Staubli VAL3: Action.pjx

--- Action.pjx ---
Parameters version=s8.10.3Cs9_BS2093 stackSize=5000 millimeterUnit=true
Program file=_tActCtrl.pgx
Program file=action.pgx
Program file=action_do.pgx
Program file=addActCmd.pgx
Program file=checkMoveId.pgx
Program file=clearActStack.pgx
Program file=create.pgx
Program file=init.pgx
Program file=kill.pgx
Program file=moveJToJoint.pgx
Program file=moveLJToPoint.pgx
Program file=pushActCmd.pgx
Program file=removeActCmd.pgx
Program file=resetMoveId.pgx
Program file=start.pgx
Program file=stop.pgx
Data file=Action.dtx
Library alias=io path=Disk://source/projectSource/io/io.pjx
Library alias=rs path=Disk://source/projectSource/robotStatus/robotStatus.pjx
Library alias=actionData path=Disk://data/actionData/actionData.pjx
Type name=actionIO path=Disk://source/template/action/action.pjx
Type name=actCmdType path=Disk://source/template/actCmd/actCmd.pjx

--- Action.dtx ---
actCmdType actCmd[40]
  [0]
    bool bActFinish
    num nActionID
    num nMoveID
    string sActName
  [1]
    bool bActFinish
    num nActionID
    num nMoveID
    string sActName
  [2]
    bool bActFinish
    num nActionID
    num nMoveID
    string sActName
  [3]
    bool bActFinish
    num nActionID
    num nMoveID
    string sActName
  [4]
    bool bActFinish
    num nActionID
    num nMoveID
    string sActName
  [5]
    bool bActFinish
    num nActionID
    num nMoveID
    string sActName
  [6]
    bool bActFinish
    num nActionID
    num nMoveID
    string sActName
  [7]
    bool bActFinish
    num nActionID
    num nMoveID
    string sActName
  [8]
    bool bActFinish
    num nActionID
    num nMoveID
    string sActName
  [9]
    bool bActFinish
    num nActionID
    num nMoveID
    string sActName
  [10]
    bool bActFinish
    num nActionID
    num nMoveID
    string sActName
  [11]
    bool bActFinish
    num nActionID
    num nMoveID
    string sActName
  [12]
    bool bActFinish
    num nActionID
    num nMoveID
    string sActName
  [13]
    bool bActFinish
    num nActionID
    num nMoveID
    string sActName
  [14]
    bool bActFinish
    num nActionID
    num nMoveID
    string sActName
  [15]
    bool bActFinish
    num nActionID
    num nMoveID
    string sActName
  [16]
    bool bActFinish
    num nActionID
    num nMoveID
    string sActName
  [17]
    bool bActFinish
    num nActionID
    num nMoveID
    string sActName
  [18]
    bool bActFinish
    num nActionID
    num nMoveID
    string sActName
  [19]
    bool bActFinish
    num nActionID
    num nMoveID
    string sActName
  [20]
    bool bActFinish
    num nActionID
    num nMoveID
    string sActName
  [21]
    bool bActFinish
    num nActionID
    num nMoveID
    string sActName
  [22]
    bool bActFinish
    num nActionID
    num nMoveID
    string sActName
  [23]
    bool bActFinish
    num nActionID
    num nMoveID
    string sActName
  [24]
    bool bActFinish
    num nActionID
    num nMoveID
    string sActName
  [25]
    bool bActFinish
    num nActionID
    num nMoveID
    string sActName
  [26]
    bool bActFinish
    num nActionID
    num nMoveID
    string sActName
  [27]
    bool bActFinish
    num nActionID
    num nMoveID
    string sActName
  [28]
    bool bActFinish
    num nActionID
    num nMoveID
    string sActName
  [29]
    bool bActFinish
    num nActionID
    num nMoveID
    string sActName
  [30]
    bool bActFinish
    num nActionID
    num nMoveID
    string sActName
  [31]
    bool bActFinish
    num nActionID
    num nMoveID
    string sActName
  [32]
    bool bActFinish
    num nActionID
    num nMoveID
    string sActName
  [33]
    bool bActFinish
    num nActionID
    num nMoveID
    string sActName
  [34]
    bool bActFinish
    num nActionID
    num nMoveID
    string sActName
  [35]
    bool bActFinish
    num nActionID
    num nMoveID
    string sActName
  [36]
    bool bActFinish
    num nActionID
    num nMoveID
    string sActName
  [37]
    bool bActFinish
    num nActionID
    num nMoveID
    string sActName
  [38]
    bool bActFinish
    num nActionID
    num nMoveID
    string sActName
  [39]
    bool bActFinish
    num nActionID
    num nMoveID
    string sActName
actionIO aActionUsing
  [0]
    num nActIO
    num nActResult
    num nActType
actionIO actPrt[40]
  [0]
    num nActIO
    num nActResult
    num nActType
  [1]
    num nActIO
    num nActResult
    num nActType
  [2]
    num nActIO
    num nActResult
    num nActType
  [3]
    num nActIO
    num nActResult
    num nActType
  [4]
    num nActIO
    num nActResult
    num nActType
  [5]
    num nActIO
    num nActResult
    num nActType
  [6]
    num nActIO
    num nActResult
    num nActType
  [7]
    num nActIO
    num nActResult
    num nActType
  [8]
    num nActIO
    num nActResult
    num nActType
  [9]
    num nActIO
    num nActResult
    num nActType
  [10]
    num nActIO
    num nActResult
    num nActType
  [11]
    num nActIO
    num nActResult
    num nActType
  [12]
    num nActIO
    num nActResult
    num nActType
  [13]
    num nActIO
    num nActResult
    num nActType
  [14]
    num nActIO
    num nActResult
    num nActType
  [15]
    num nActIO
    num nActResult
    num nActType
  [16]
    num nActIO
    num nActResult
    num nActType
  [17]
    num nActIO
    num nActResult
    num nActType
  [18]
    num nActIO
    num nActResult
    num nActType
  [19]
    num nActIO
    num nActResult
    num nActType
  [20]
    num nActIO
    num nActResult
    num nActType
  [21]
    num nActIO
    num nActResult
    num nActType
  [22]
    num nActIO
    num nActResult
    num nActType
  [23]
    num nActIO
    num nActResult
    num nActType
  [24]
    num nActIO
    num nActResult
    num nActType
  [25]
    num nActIO
    num nActResult
    num nActType
  [26]
    num nActIO
    num nActResult
    num nActType
  [27]
    num nActIO
    num nActResult
    num nActType
  [28]
    num nActIO
    num nActResult
    num nActType
  [29]
    num nActIO
    num nActResult
    num nActType
  [30]
    num nActIO
    num nActResult
    num nActType
  [31]
    num nActIO
    num nActResult
    num nActType
  [32]
    num nActIO
    num nActResult
    num nActType
  [33]
    num nActIO
    num nActResult
    num nActType
  [34]
    num nActIO
    num nActResult
    num nActType
  [35]
    num nActIO
    num nActResult
    num nActType
  [36]
    num nActIO
    num nActResult
    num nActType
  [37]
    num nActIO
    num nActResult
    num nActType
  [38]
    num nActIO
    num nActResult
    num nActType
  [39]
    num nActIO
    num nActResult
    num nActType
bool bPushToStack
public num _nActStackIndex
num _nNextId
public num _nPuleStartClk[128]
public num nMoveIDRef
num nMoveIdMax = 100
num nSyncMoveID

--- start.pgx ---
program start()
begin
end

--- _tActCtrl.pgx ---
program _tActCtrl()
  local num l_n
  local num l_nMoveID
  local num l_nDeltaMoveId
begin
  do
    for l_n=0 to size(actCmd)-1
      //当moveID有值且没有将动作放入动作堆栈时：
      if actCmd[l_n].nMoveID>=0 and bPushToStack==false
        l_nMoveID=getMoveId()
        if l_nMoveID<nMoveIdMax*0.2 and actCmd[l_n].nMoveID>nMoveIdMax*0.8
          // l_nMoveID roll over
          l_nDeltaMoveId=(l_nMoveID+nMoveIdMax)-actCmd[l_n].nMoveID
        elseIf l_nMoveID>nMoveIdMax*0.8 and actCmd[l_n].nMoveID<nMoveIdMax*0.2
          // actCmd[l_n].nMoveID roll over
          l_nDeltaMoveId=l_nMoveID-(actCmd[l_n].nMoveID+nMoveIdMax)
        else
          //normal condition
          l_nDeltaMoveId=(l_nMoveID-actCmd[l_n].nMoveID)
        endIf

        if l_nDeltaMoveId>1 and actPrt[l_n].nActType!=2
          // action control error, set alarm
          call rs:setAlarm(209,l_nDeltaMoveId)
        elseIf l_nDeltaMoveId>=0
          if actCmd[l_n].nActionID>=0
            //execute cmd
            call action(actCmd[l_n].nActionID,actCmd[l_n].bActFinish)
            if actCmd[l_n].bActFinish[0]
              // action done,remove cmd
              call removeActCmd(l_n)
            endIf
          else
            //动作的范围超限
            call rs:setAlarm(208,actCmd[l_n].nActionID)
          endIf
        endIf
      endIf
    endFor
    delay(0)
  until false
end

--- action.pgx ---
program action(num x_nActID, bool& x_bFinish[])
  local bool l_bErr
  local num l_n
  local num l_nActIO
  local num l_nActRslt
  local num l_nActType
begin
  //类型nType      结果nResult 含义如下     l_nActIO
  //	1=out	       0=false 1=true          IO的索引号
  //	2=Pulse	     l_nActRslt 延时n s      IO的索引号

  if x_nActID>=0 and x_nActID<size(actCmd)
    //execute action group x_nActID
    l_n=0
    if x_bFinish[l_n]==false
      l_nActIO=actPrt[x_nActID].nActIO[l_n]
      l_nActType=actPrt[x_nActID].nActType[l_n]
      l_nActRslt=actPrt[x_nActID].nActResult[l_n]
      //
      if l_nActIO>=0
        switch l_nActType
          case 1
            //set output
            if l_nActRslt==0
              call io:setDigOutput(io:dOutput[l_nActIO],false,l_bErr)
            elseIf l_nActRslt==1
              call io:setDigOutput(io:dOutput[l_nActIO],true,l_bErr)
            endIf
            x_bFinish[l_n]=true
          break

          case 2
            //pulse ouput
            if l_nActRslt>0
              if _nPuleStartClk[l_nActIO]<0
                call io:setDigOutput(io:dOutput[l_nActIO],true,l_bErr)
                _nPuleStartClk[l_nActIO]=clock()
              else
                if clock()-_nPuleStartClk[l_nActIO]>l_nActRslt
                  call io:setDigOutput(io:dOutput[l_nActIO],false,l_bErr)
                  _nPuleStartClk[l_nActIO]=-1
                  x_bFinish[l_n]=true
                endIf
              endIf
            endIf
          break

        endSwitch
      else
        //none
        x_bFinish[l_n]=true
      endIf
    endIf
  endIf
end

--- action_do.pgx ---
public program action_do(num x_nIndex)
  local num l_nType
  local string l_sType
  local bool l_bActive
  local string l_sBoolValue
  local num l_nBoolValue
  local num l_nIOindex
  local num l_nPulseValue
  local num l_i
begin
  for l_i = 0 to size(actionData:aActItem[x_nIndex].aActItem)-1
    l_sType=actionData:aActItem[x_nIndex].aActItem[l_i].sIOtype
    l_bActive=(actionData:aActItem[x_nIndex].aActItem[l_i].bActive==true)
    l_sBoolValue=actionData:aActItem[x_nIndex].aActItem[l_i].sValue
    l_nIOindex=actionData:aActItem[x_nIndex].aActItem[l_i].nIOindex
    l_nPulseValue=actionData:aActItem[x_nIndex].aActItem[l_i].nPulseValue
    switch l_sBoolValue
      case "ON"
        l_nBoolValue=1
      break
      case "OFF"
        l_nBoolValue=0
      break
    endSwitch
    if l_bActive
      switch l_sType
        case "IN"
          call addActCmd(1,3,l_nIOindex,l_nBoolValue)
        break
        case "OUT"
          call addActCmd(1,1,l_nIOindex,l_nBoolValue)
        break
        case "PULSE"
          call addActCmd(1,2,l_nIOindex,l_nPulseValue)
        break

      endSwitch
    endIf
  endFor
  popUpMsg("执行动作："+toString("",x_nIndex))
end

--- addActCmd.pgx ---
public program addActCmd(num x_nPercent, num x_nInOutType, num x_nInOutIndex, num x_nInOutValue)
// //作用：将动作添加到动作堆栈中
//   //用法：x_nPercent 指的是运动的百分比，其值为0到1，如该值为0.8，
//   则代表一条运动指令运动到80%时，执行该动作。
//   //x_nInOutType指的是输入输出的类型  1代表输出Out  2代表脉冲Pulse 3代表输入In
//   //x_nInOutIndex是输入或者输出的索引号，默认值为0到95
//   //x_nInOutValue 指的是输入输出或者脉冲的值
//   //类型x_nInOutType        结果x_nInOutValue
//   // 1=out                0=false 1=true
//   // 2=Pulse              延时x_nInOutValue秒后信号置为OFF.
//   // 3=in                0=false  1=true
// 
//   //示例： call addActCmd(0.8,1,32,1)   代表一条运行指令运动到80%时，输出io库中的第32号信号dOutput为ON
//   //      call addActCmd(0.7,2,33,2.2) 代表一条运行指令运动到70%时，脉冲输出io库中的第33号信号dOutput为ON，然后2.2秒后将该信号置位OFF.
//   //      call addActCmd(0.6,3,34,1)   代表一条运行指令运动到60%时,等待输入io库中的第33号信号为ON，注意：该信号如果不满足则会阻塞运动任务
  local bool l_bErr
begin
  //作用：将动作添加到动作堆栈中，动作包含输出信号、脉冲信号及等待信号
  //用法：
  //x_nPercent 指的是运动的百分比，其值为0到1，如该值为0.8，则代表一条运动指令运动到80%时，执行该动作。
  //x_nInOutType指的是输入输出的类型  1代表输出Out	 2代表脉冲Pulse	3代表输入In
  //x_nInOutIndex是输入或者输出的索引号，默认值为0到95
  //x_nInOutValue 指的是输入输出或者脉冲的值
  //类型x_nInOutType        结果x_nInOutValue
  //	1=out	               0=false 1=true
  //	2=Pulse	             延时x_nInOutValue秒后信号置为OFF.
  //	3=in	               0=false  1=true
  //示例： call addActCmd(0.8,1,32,1)   代表一条运行指令运动到80%时，输出io库中的第32号信号dOutput为ON
  //      call addActCmd(0.7,2,33,2.2) 代表一条运行指令运动到70%时，脉冲输出io库中的第33号信号dOutput为ON，然后2.2秒后将该信号置位OFF.
  //      call addActCmd(0.6,3,34,1)   代表一条运行指令运动到60%时,等待输入io库中的第33号信号为ON，注意：该信号如果不满足则会阻塞运动任务

  //nMoveIDRef: 运动的MoveID，通过movel或者movej获得。

  if x_nPercent>1 or x_nPercent<0
    //动作的百分比要正确
    call rs:setAlarm(202,x_nPercent)
  elseIf !(x_nInOutType==1 or x_nInOutType==2 or x_nInOutType==3)
    //动作的输入输出的类型要正确
    call rs:setAlarm(203,x_nInOutType)
  elseIf x_nInOutIndex<32 or x_nInOutIndex>io:nMaxdigital-1
    //索引号的范围是32到95
    call rs:setAlarm(204,x_nInOutIndex)
  else
    //OUT输出的动作放入到动作堆栈
    switch x_nInOutType
      case 1,2
        //判断OUT的x_nInOutValue范围
        if x_nInOutType==1 and !(x_nInOutValue==0 or x_nInOutValue==1)
          call rs:setAlarm(205,x_nInOutValue)
        elseIf x_nInOutType==2 and  x_nInOutValue<0
          call rs:setAlarm(206,x_nInOutValue)
        endIf
        aActionUsing.nActType=x_nInOutType
        aActionUsing.nActIO=x_nInOutIndex
        aActionUsing.nActResult=x_nInOutValue
        call pushActCmd(nMoveIDRef+x_nPercent,aActionUsing)
        if x_nPercent==1
          waitEndMove()
        endIf
      break
      case 3
        //IN输入动作，运动任务会等待该信号，即该信号会阻塞该运动任务

        if x_nPercent==1
          waitEndMove()
        else
          wait(getMoveId()>=nMoveIDRef+x_nPercent)
        endIf
        if x_nInOutValue==0
          call io:waitDigInput(io:dInput[x_nInOutIndex],false,l_bErr)
        elseIf x_nInOutValue==1
          call io:waitDigInput(io:dInput[x_nInOutIndex],true,l_bErr)
        else
          call rs:setAlarm(207,x_nInOutValue)
        endIf
      break
    endSwitch
  endIf

end

--- checkMoveId.pgx ---
program checkMoveId()
begin
  //作用：检查当前的moveiD,当前的MoveID到达设置的最大值时，设置MoveID为0，避免MoveID编程随机值。
  _nNextId=nextMoveId()
  if _nNextId>nMoveIdMax
    call rs:setAlarm(210,_nNextId)
  elseIf _nNextId==nMoveIdMax
    wait(getMoveId()>=nMoveIDRef+nSyncMoveID)
    setMoveId(0)
  else
    //2.正常的值
    wait(getMoveId()>=nMoveIDRef+nSyncMoveID)
  endIf

end

--- clearActStack.pgx ---
public program clearActStack()
  local num l_n
begin
  for l_n=0 to size(_nPuleStartClk)-1
    _nPuleStartClk[l_n]=-1
  endFor
  _nActStackIndex=0
  for l_n=0 to size(actCmd)-1
    call removeActCmd(l_n)
  endFor
end

--- create.pgx ---
public program create()
begin
  call init()
  //action control management
  taskKill("actCtrl")
  taskCreate "actCtrl",100,_tActCtrl()
  wait(taskStatus("actCtrl")==1)
end

--- init.pgx ---
public program init()
begin
  //更改_nPuleStartClk的大小
  if size(_nPuleStartClk)!=io:nMaxdigital
    resize(_nPuleStartClk,1,io:nMaxdigital)
    libSave()
  endIf
  //num
  _nActStackIndex=0
  //Bool
  bPushToStack=false
  //
  call clearActStack()
  //
  setMoveId(0)
end

--- kill.pgx ---
public program kill()
begin
  //Kill Task
  taskKill("actCtrl")
  wait(taskStatus("actCtrl")==-1)
  call clearActStack()
end

--- moveJToJoint.pgx ---
public program moveJToJoint(joint x_jTarget, tool x_tTool, mdesc x_mSpeed)
// //作用：用关节运动的方式移动到目标点。
//   //参数：
//   //x_jTarget: 目标点Joint值
//   //  x_tTool：去目标点使用的工具值
//   //  x_mSpeed:去目标点使用的速度值
//   //x_bWaitEndmove:到达目标点，没有混合，为true则是严格到达目标点
  local bool l_bInRange
begin
  //作用：用关节运动的方式移动到目标点。
  //参数：
  //x_jTarget: 目标点Joint值
  //  x_tTool：去目标点使用的工具值
  //  x_mSpeed:去目标点使用的速度值
  //  x_bWaitEndmove:到达目标点，没有混合，为true则是严格到达目标点

  l_bInRange=isInRange(x_jTarget)
  if l_bInRange==true
    nMoveIDRef=movej(x_jTarget,x_tTool,x_mSpeed)
    call checkMoveId()
  else
    //超出机器人限位
    call rs:setAlarm(221,-1)
  endIf

end

--- moveLJToPoint.pgx ---
public program moveLJToPoint(bool x_bMoveL, point x_pPoint, tool x_tTool, mdesc x_mSpeed)
// //作用：用直线或者关节运动的方式移动到目标Point点。
//   //参数：
//   //x_bMoveL: 为true时，直线运动到该点；为false时，关节运动到该Point点
//   //x_pPoint:目标点Point值
//   // x_tTool：去目标点使用的工具值
//   //x_bReference: 将点位转换为Joint来判断改为是否超限位，当该值为true时，使用jHome作为参考，为falses时，使用当前的关节值。
//   // x_mSpeed:去目标点使用的速度值
//    //x_bWaitEndmove:到达目标点，没有混合，为true则是严格到达目标点
//   //示例  call moveLJToPoint(true,data:pPointRx[0],data:tTool[0],false,data:mMdesc[0])
  local bool l_bResult
  local joint l_jHere
  local bool l_bInRange
  local jointRx l_jTarget
begin
  //作用：用直线或者关节运动的方式移动到目标Point点。
  //参数：
  //x_bMoveL: 为true时，直线运动到该点；为false时，关节运动到该Point点
  //x_pPoint:目标点Point值
  // x_tTool：去目标点使用的工具值
  //x_bReference: 将点位转换为Joint来判断改为是否超限位，当该值为true时，使用jHome作为参考，为false时，使用当前的关节值。
  // x_mSpeed:去目标点使用的速度值
  // x_bWaitEndmove:到达目标点，没有混合，为true则是严格到达目标点
  //示例  call moveLJToPoint(true,data:pPointRx[0],data:tTool[0],false,data:mMdesc[0])
  l_jHere=herej()
  l_bResult=pointToJoint(x_tTool,l_jHere,x_pPoint,l_jTarget)

  //check in range
  if l_bResult
    l_bInRange=isInRange(l_jTarget)
  else
    l_bInRange=false
  endIf

  if l_bInRange==true
    if x_bMoveL==true
      nMoveIDRef=movel(x_pPoint,x_tTool,x_mSpeed)
    else
      nMoveIDRef=movej(x_pPoint,x_tTool,x_mSpeed)
    endIf
    call checkMoveId()
  else
    //超出机器人限位
    call rs:setAlarm(220,-1)
  endIf

end

--- pushActCmd.pgx ---
program pushActCmd(num x_nMoveID, actionIO x_actPrt)
begin
  //add to action stack, excute act command in actCtrl task, to optmize cycle time
  setMutex(bPushToStack)
  _nActStackIndex=(_nActStackIndex+1)%size(actCmd)
  if actCmd[_nActStackIndex].nMoveID<0
    actCmd[_nActStackIndex].nMoveID=x_nMoveID
    actCmd[_nActStackIndex].nActionID =_nActStackIndex
    actPrt[_nActStackIndex]=x_actPrt
  else
    call rs:setAlarm(201,-1)
  endIf
  bPushToStack=false
end

--- removeActCmd.pgx ---
program removeActCmd(num x_nStackIndex)
begin
  actCmd[x_nStackIndex].nMoveID=-1
  actCmd[x_nStackIndex].nActionID=-1
  actCmd[x_nStackIndex].bActFinish[0]=false
end

--- resetMoveId.pgx ---
public program resetMoveId()
  local num l_nNextId
begin
  //reset move id to avoid move id overflow
  l_nNextId=nextMoveId()
  if l_nNextId>=nMoveIdMax
    setMoveId(0)
  endIf
end

--- stop.pgx ---
program stop()
begin
end
